(* IEC 61131-3 sources: codesys-framework/txt/application/ToDo/Utils/FB_Timer, 4 files *)

(* ---- GetTime.method.st ---- *)
METHOD GetTime : TIME
VAR_INPUT
END_VAR

// --- BEGIN IMPLEMENTATION ---

GetTime := _tTotal;

(* ---- Reset.method.st ---- *)
METHOD Reset
VAR_INPUT
END_VAR

// --- BEGIN IMPLEMENTATION ---

_tStart := TO_TIME(SysTimeGetMs());
_tEnd := TO_TIME(SysTimeGetMs());
_tDelta := T#0MS;
_tPrevious := T#0MS;
_tTotal := T#0MS;

(* ---- Start.method.st ---- *)
METHOD Start
VAR_INPUT
END_VAR

// --- BEGIN IMPLEMENTATION ---

_xOn := TRUE;

(* ---- Stop.method.st ---- *)
METHOD Stop
VAR_INPUT
END_VAR

// --- BEGIN IMPLEMENTATION ---

_xOn := FALSE;
